(* Logix 5000 project; controller TFF vendor 1 type 14 code 107 rev 34.11; software revision 34.03; part 33 of 36 *)
(* tags used below, declared in another part *)
   Address : DINT;   // Temp Address
   Index : DINT;   // Index
   FlowPath : FlowPath[64];   // Flow Path Array
   PipeAnimation : PipeAnimation;   // HMI Pipe Animation Array
   PipeStatValueHMI : INT[224];   // Pipe Animation Value For HMI
   Rack_Murr_Node0_Smart : IO_Station;   // Status of Node 0 Smart
   Rack_Murr_Node1_TF2S : IO_Station;   // Status of Node 1 TF2S
   Rack_Murr_Node1_TF3S : IO_Station;   // Status of Node 1 TF3S
   Rack_Murr_Node3_PUMP : IO_Station;   // Status of Node 3 Pump
   Rack_Murr_Node4_Instrum_TFF1 : IO_Station;   // Status of Node 4 Instrum TFF1
   Rack_Murr_Node4_Instrum_TFF2 : IO_Station;   // Status of Node 4 Instrum TFF2
   Rack_Murr_Node4_Instrum_TFF3 : IO_Station;   // Status of Node 4 Instrum TFF3
   Rack_Murr_Node4_Instrum_TFF4 : IO_Station;   // Status of Node 4 Instrum TFF4
   Rack_Murr_Node4_Instrum_TFF5 : IO_Station;   // Status of Node 4 Instrum TFF5
   Rack_Murr_Node5_Tank100 : IO_Station;   // Status of Node 5 Tank 100L
   Rack_Murr_Node5_Tank250 : IO_Station;   // Status of Node 5 Tank 250L
   Rack_Murr_Node5_Tank50 : IO_Station;   // Status of Node 5 Tank 50L
   Rack_Murr_Node6_IND331_WI001 : IO_Station;   // Status of Node 6 IND331 WI001
   Rack_Murr_Node7_IND131_WI101 : IO_Station;   // Status of Node 7 IND131 WI101
   SIC001 : ALIAS FOR Drive[1];   // Feed Pump
   SIC002 : ALIAS FOR Drive[2];   // Transfer Pump
   Tank : TankManagement;   // Tank Management
   WI001 : ALIAS FOR AnalogPoint[15];   // Feed Bag Weight
   WI101 : ALIAS FOR AnalogPoint[0];   // Filtrate Weight
(* Process, continued *)

ROUTINE PipeAnimationHMI   (* ladder *)
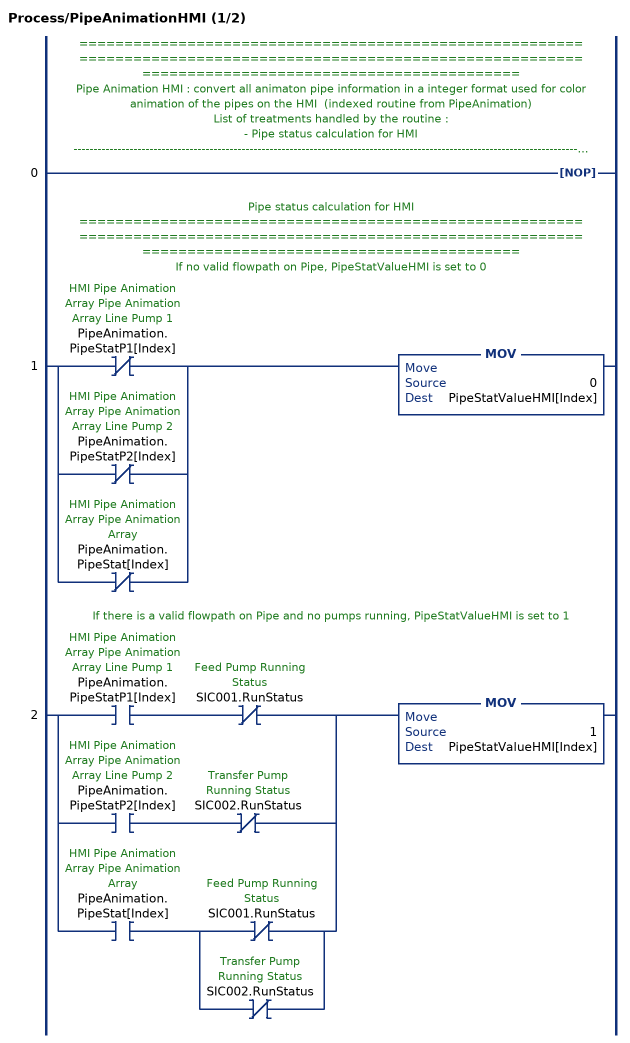
   // ==========================================================================================================================================================
   //                          Pipe Animation HMI : convert all animaton pipe information in a integer format used for color animation of the pipes on the HMI  (indexed routine from PipeAnimation)
   //                                                     List of treatments handled by the routine :
   //                                                          - Pipe status calculation for HMI
   //                                                     -----------------------------------------------------------------------------------------------------------------------------------------------------
   //                                                     History
   //                                                          2019-AUG-13 - Actemium - B. Roch - Initial version for Candidate Release 3.00.00.00.a
   // ========================================================================================================================================================
   0: NOP();
   // Pipe status calculation for HMI
   // ==========================================================================================================================================================
   // If no valid flowpath on Pipe, PipeStatValueHMI is set to 0
   1: [XIO(PipeAnimation.PipeStatP1[Index]) ,XIO(PipeAnimation.PipeStatP2[Index]) ,XIO(PipeAnimation.PipeStat[Index]) ]MOV(0,PipeStatValueHMI[Index]);
   // If there is a valid flowpath on Pipe and no pumps running, PipeStatValueHMI is set to 1
   2: [XIC(PipeAnimation.PipeStatP1[Index]) XIO(SIC001.RunStatus) ,XIC(PipeAnimation.PipeStatP2[Index]) XIO(SIC002.RunStatus) ,XIC(PipeAnimation.PipeStat[Index]) [XIO(SIC001.RunStatus) ,XIO(SIC002.RunStatus) ] ]MOV(1,PipeStatValueHMI[Index]);
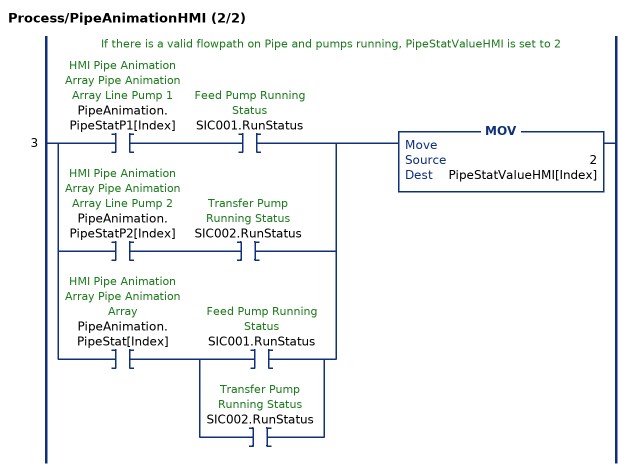
   // If there is a valid flowpath on Pipe and pumps running, PipeStatValueHMI is set to 2
   3: [XIC(PipeAnimation.PipeStatP1[Index]) XIC(SIC001.RunStatus) ,XIC(PipeAnimation.PipeStatP2[Index]) XIC(SIC002.RunStatus) ,XIC(PipeAnimation.PipeStat[Index]) [XIC(SIC001.RunStatus) ,XIC(SIC002.RunStatus) ] ]MOV(2,PipeStatValueHMI[Index]);
END_ROUTINE

ROUTINE Scale   (* function block diagram *)
// Scale Routine
   SHEET 1
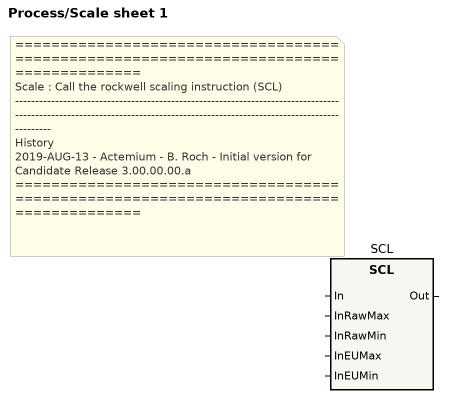
   // ======================================================================================
   // Scale : Call the rockwell scaling instruction (SCL)
   // ------------------------------------------------------------------------------------------------------------------------------------------------------------------
   // ---------
   // History
   //    2019-AUG-13 - Actemium - B. Roch - Initial version for Candidate Release 3.00.00.00.a
   // ======================================================================================
   SCL : SCL();   // unwired pins: In InRawMax InRawMin InEUMax InEUMin Out
END_ROUTINE

ROUTINE Station_Status   (* ladder *)
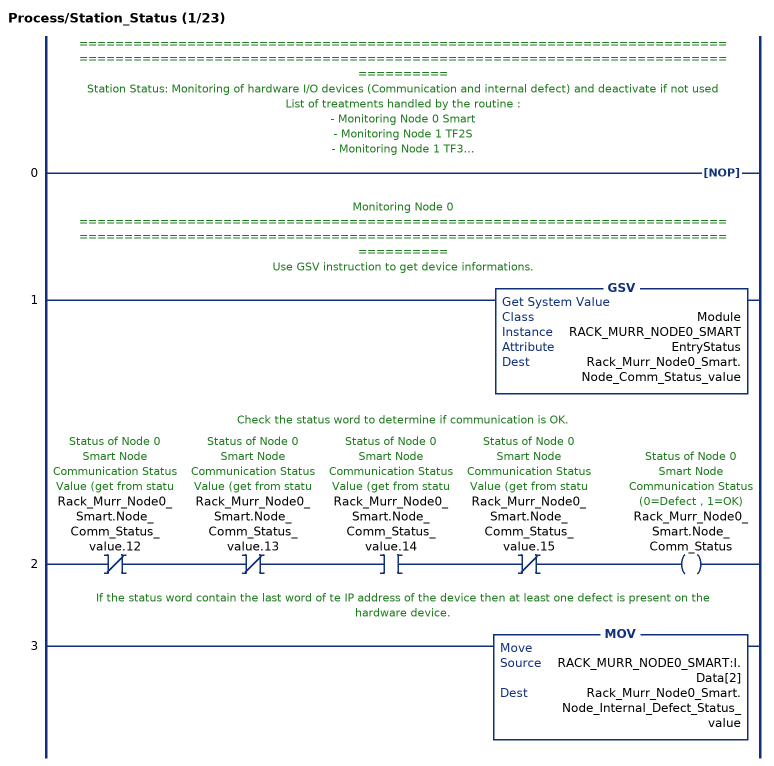
   // ==========================================================================================================================================================
   //                                                                   Station Status: Monitoring of hardware I/O devices (Communication and internal defect) and deactivate if not used
   //                                                     List of treatments handled by the routine :
   //                                                        - Monitoring Node 0 Smart
   //                                                        - Monitoring Node 1 TF2S
   //                                                        - Monitoring Node 1 TF3S
   //                                                        - Monitoring Node 3 PUMP
   //                                                        - Monitoring Node 4 INTRUM TFF1
   //                                                        - Monitoring Node 4 INTRUM TFF2
   //                                                        - Monitoring Node 4 INTRUM TFF3
   //                                                        - Monitoring Node 4 INTRUM TFF4
   //                                                        - Monitoring Node 4 INTRUM TFF5
   //                                                        - Monitoring Node 5 TANK50
   //                                                        - Monitoring Node 5 TANK100
   //                                                        - Monitoring Node 5 TANK250
   //                                                        - Monitoring Node 6 IND331 WI001
   //                                                        - Monitoring Node 7 IND131 WI101
   //                                                        - Deactivate / Activate devices
   //                                                     -----------------------------------------------------------------------------------------------------------------------------------------------------
   //                                                     History
   //                                                          2019-AUG-13 - Actemium - B. Roch - Initial version for Candidate Release 3.00.00.00.a
   // ========================================================================================================================================================
   0: NOP();
   // Monitoring Node 0
   // ==========================================================================================================================================================
   // Use GSV instruction to get device informations.
   1: GSV(Module,RACK_MURR_NODE0_SMART,EntryStatus,Rack_Murr_Node0_Smart.Node_Comm_Status_value);
   // Check the status word to determine if communication is OK.
   2: XIO(Rack_Murr_Node0_Smart.Node_Comm_Status_value.12)XIO(Rack_Murr_Node0_Smart.Node_Comm_Status_value.13)XIC(Rack_Murr_Node0_Smart.Node_Comm_Status_value.14)XIO(Rack_Murr_Node0_Smart.Node_Comm_Status_value.15)OTE(Rack_Murr_Node0_Smart.Node_Comm_Status);
   // If the status word contain the last word of te IP address of the device then at least one defect is present on the hardware device.
   3: MOV(RACK_MURR_NODE0_SMART:I.Data[2],Rack_Murr_Node0_Smart.Node_Internal_Defect_Status_value);
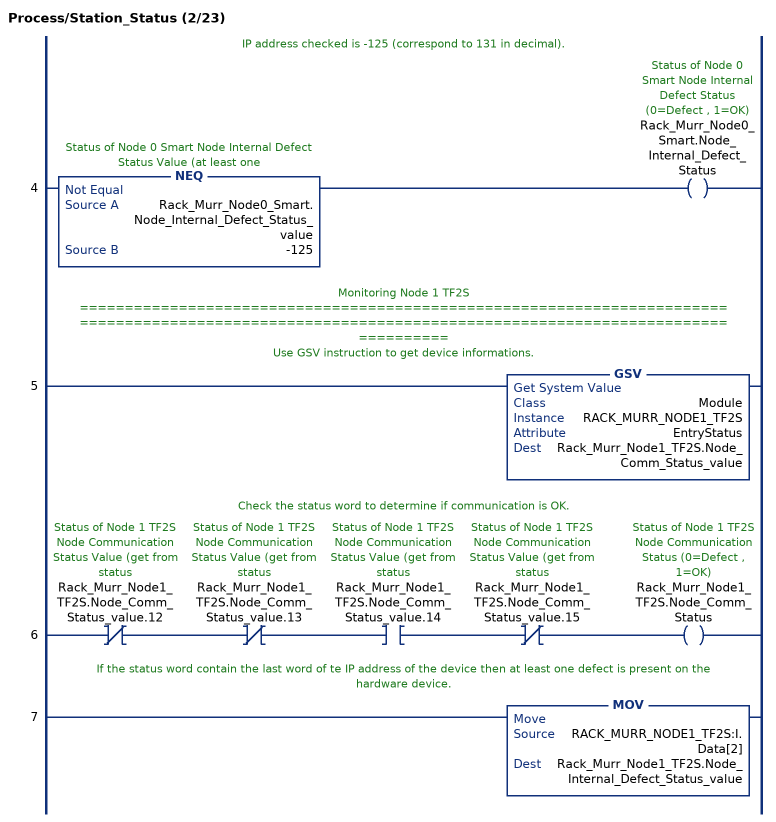
   // IP address checked is -125 (correspond to 131 in decimal).
   4: NEQ(Rack_Murr_Node0_Smart.Node_Internal_Defect_Status_value,-125)OTE(Rack_Murr_Node0_Smart.Node_Internal_Defect_Status);
   // Monitoring Node 1 TF2S
   // ==========================================================================================================================================================
   // Use GSV instruction to get device informations.
   5: GSV(Module,RACK_MURR_NODE1_TF2S,EntryStatus,Rack_Murr_Node1_TF2S.Node_Comm_Status_value);
   // Check the status word to determine if communication is OK.
   6: XIO(Rack_Murr_Node1_TF2S.Node_Comm_Status_value.12)XIO(Rack_Murr_Node1_TF2S.Node_Comm_Status_value.13)XIC(Rack_Murr_Node1_TF2S.Node_Comm_Status_value.14)XIO(Rack_Murr_Node1_TF2S.Node_Comm_Status_value.15)OTE(Rack_Murr_Node1_TF2S.Node_Comm_Status);
   // If the status word contain the last word of te IP address of the device then at least one defect is present on the hardware device.
   7: MOV(RACK_MURR_NODE1_TF2S:I.Data[2],Rack_Murr_Node1_TF2S.Node_Internal_Defect_Status_value);
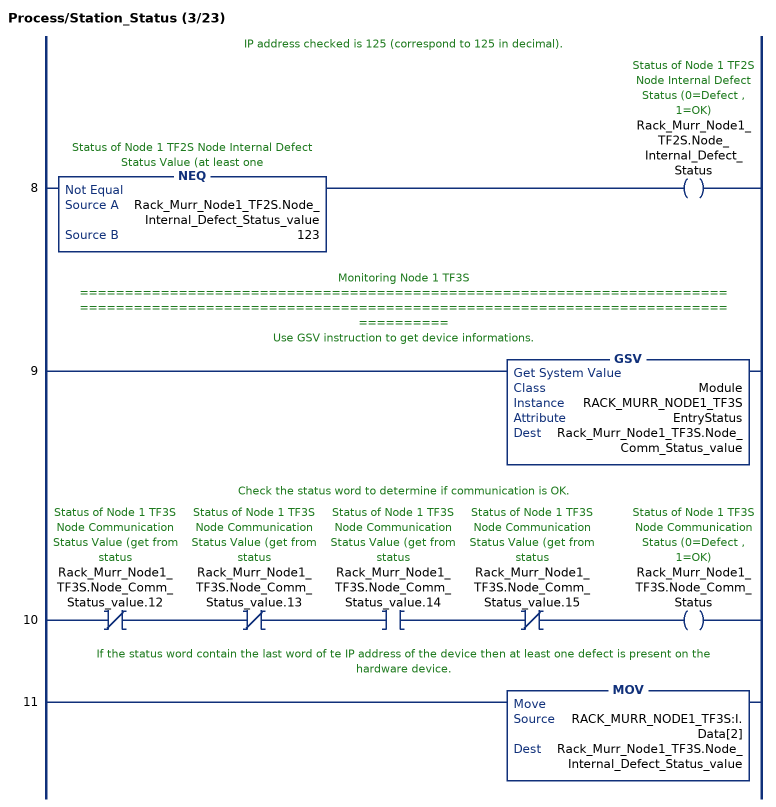
   // IP address checked is 125 (correspond to 125 in decimal).
   8: NEQ(Rack_Murr_Node1_TF2S.Node_Internal_Defect_Status_value,123)OTE(Rack_Murr_Node1_TF2S.Node_Internal_Defect_Status);
   // Monitoring Node 1 TF3S
   // ==========================================================================================================================================================
   // Use GSV instruction to get device informations.
   9: GSV(Module,RACK_MURR_NODE1_TF3S,EntryStatus,Rack_Murr_Node1_TF3S.Node_Comm_Status_value);
   // Check the status word to determine if communication is OK.
   10: XIO(Rack_Murr_Node1_TF3S.Node_Comm_Status_value.12)XIO(Rack_Murr_Node1_TF3S.Node_Comm_Status_value.13)XIC(Rack_Murr_Node1_TF3S.Node_Comm_Status_value.14)XIO(Rack_Murr_Node1_TF3S.Node_Comm_Status_value.15)OTE(Rack_Murr_Node1_TF3S.Node_Comm_Status);
   // If the status word contain the last word of te IP address of the device then at least one defect is present on the hardware device.
   11: MOV(RACK_MURR_NODE1_TF3S:I.Data[2],Rack_Murr_Node1_TF3S.Node_Internal_Defect_Status_value);
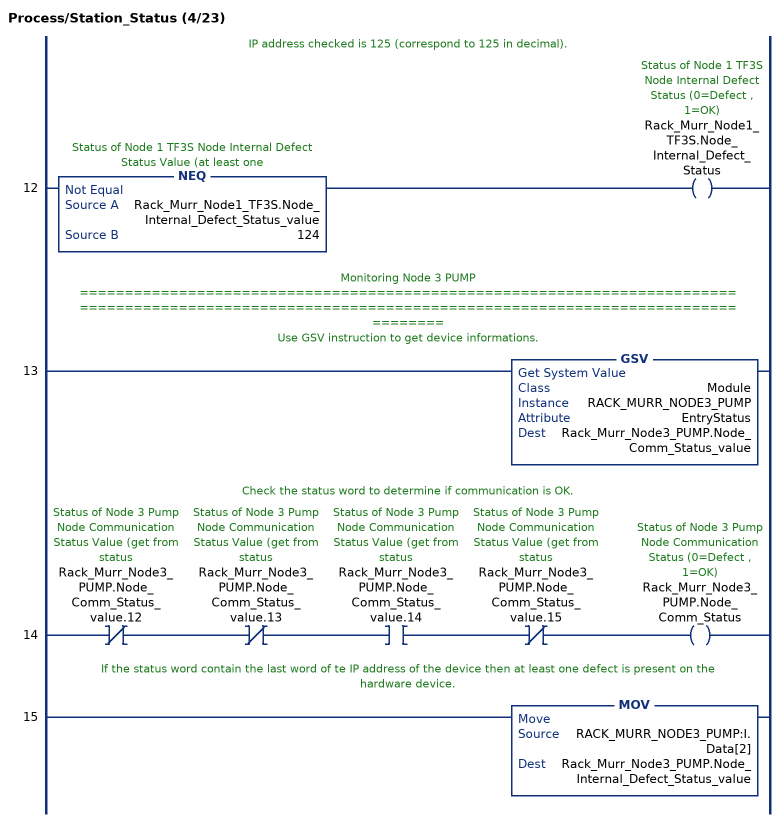
   // IP address checked is 125 (correspond to 125 in decimal).
   12: NEQ(Rack_Murr_Node1_TF3S.Node_Internal_Defect_Status_value,124)OTE(Rack_Murr_Node1_TF3S.Node_Internal_Defect_Status);
   // Monitoring Node 3 PUMP
   // ==========================================================================================================================================================
   // Use GSV instruction to get device informations.
   13: GSV(Module,RACK_MURR_NODE3_PUMP,EntryStatus,Rack_Murr_Node3_PUMP.Node_Comm_Status_value);
   // Check the status word to determine if communication is OK.
   14: XIO(Rack_Murr_Node3_PUMP.Node_Comm_Status_value.12)XIO(Rack_Murr_Node3_PUMP.Node_Comm_Status_value.13)XIC(Rack_Murr_Node3_PUMP.Node_Comm_Status_value.14)XIO(Rack_Murr_Node3_PUMP.Node_Comm_Status_value.15)OTE(Rack_Murr_Node3_PUMP.Node_Comm_Status);
   // If the status word contain the last word of te IP address of the device then at least one defect is present on the hardware device.
   15: MOV(RACK_MURR_NODE3_PUMP:I.Data[2],Rack_Murr_Node3_PUMP.Node_Internal_Defect_Status_value);
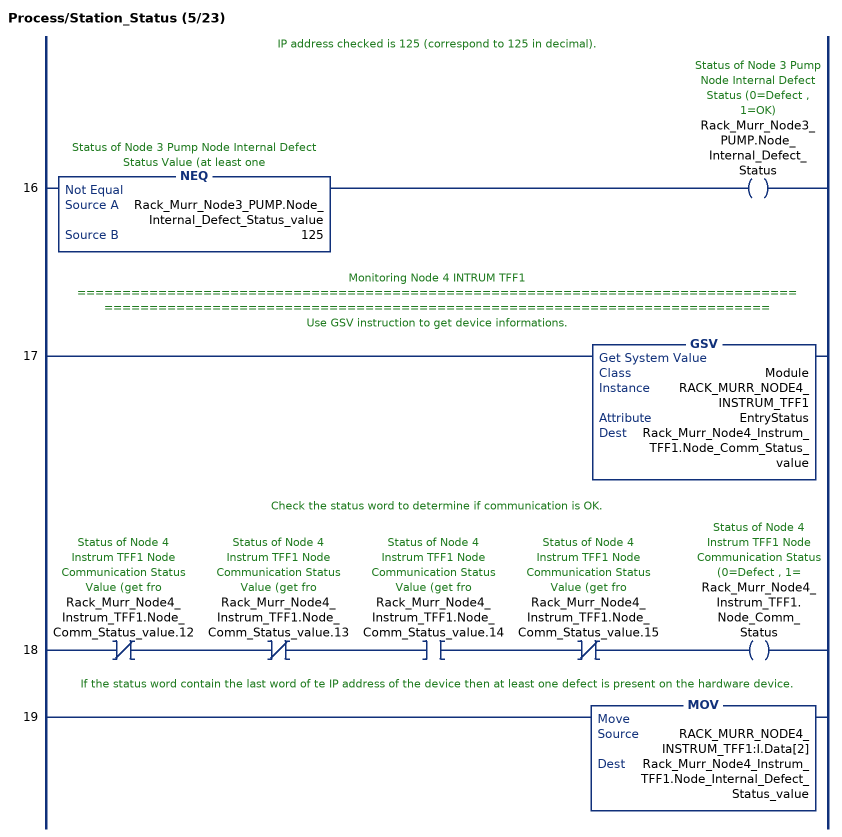
   // IP address checked is 125 (correspond to 125 in decimal).
   16: NEQ(Rack_Murr_Node3_PUMP.Node_Internal_Defect_Status_value,125)OTE(Rack_Murr_Node3_PUMP.Node_Internal_Defect_Status);
   // Monitoring Node 4 INTRUM TFF1
   // ==========================================================================================================================================================
   // Use GSV instruction to get device informations.
   17: GSV(Module,RACK_MURR_NODE4_INSTRUM_TFF1,EntryStatus,Rack_Murr_Node4_Instrum_TFF1.Node_Comm_Status_value);
   // Check the status word to determine if communication is OK.
   18: XIO(Rack_Murr_Node4_Instrum_TFF1.Node_Comm_Status_value.12)XIO(Rack_Murr_Node4_Instrum_TFF1.Node_Comm_Status_value.13)XIC(Rack_Murr_Node4_Instrum_TFF1.Node_Comm_Status_value.14)XIO(Rack_Murr_Node4_Instrum_TFF1.Node_Comm_Status_value.15)OTE(Rack_Murr_Node4_Instrum_TFF1.Node_Comm_Status);
   // If the status word contain the last word of te IP address of the device then at least one defect is present on the hardware device.
   19: MOV(RACK_MURR_NODE4_INSTRUM_TFF1:I.Data[2],Rack_Murr_Node4_Instrum_TFF1.Node_Internal_Defect_Status_value);
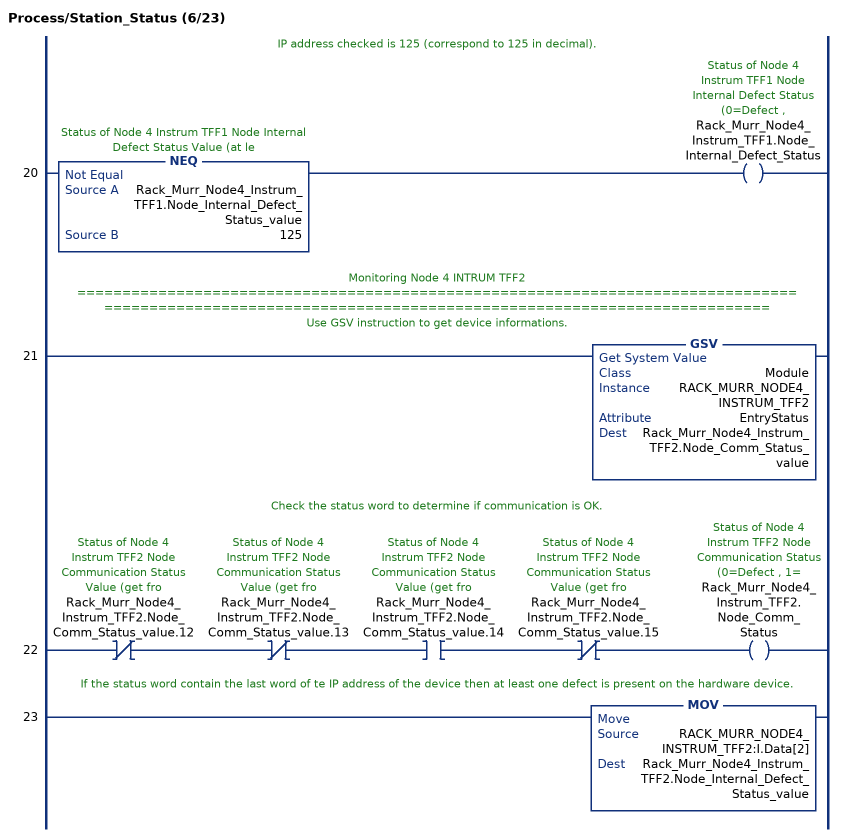
   // IP address checked is 125 (correspond to 125 in decimal).
   20: NEQ(Rack_Murr_Node4_Instrum_TFF1.Node_Internal_Defect_Status_value,125)OTE(Rack_Murr_Node4_Instrum_TFF1.Node_Internal_Defect_Status);
   // Monitoring Node 4 INTRUM TFF2
   // ==========================================================================================================================================================
   // Use GSV instruction to get device informations.
   21: GSV(Module,RACK_MURR_NODE4_INSTRUM_TFF2,EntryStatus,Rack_Murr_Node4_Instrum_TFF2.Node_Comm_Status_value);
   // Check the status word to determine if communication is OK.
   22: XIO(Rack_Murr_Node4_Instrum_TFF2.Node_Comm_Status_value.12)XIO(Rack_Murr_Node4_Instrum_TFF2.Node_Comm_Status_value.13)XIC(Rack_Murr_Node4_Instrum_TFF2.Node_Comm_Status_value.14)XIO(Rack_Murr_Node4_Instrum_TFF2.Node_Comm_Status_value.15)OTE(Rack_Murr_Node4_Instrum_TFF2.Node_Comm_Status);
   // If the status word contain the last word of te IP address of the device then at least one defect is present on the hardware device.
   23: MOV(RACK_MURR_NODE4_INSTRUM_TFF2:I.Data[2],Rack_Murr_Node4_Instrum_TFF2.Node_Internal_Defect_Status_value);
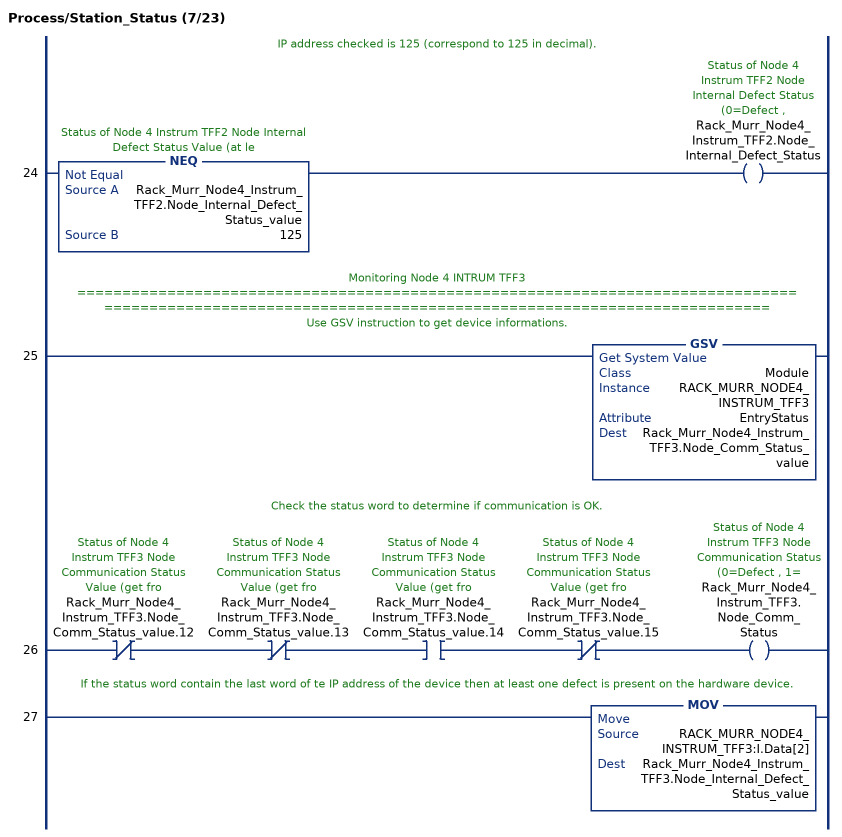
   // IP address checked is 125 (correspond to 125 in decimal).
   24: NEQ(Rack_Murr_Node4_Instrum_TFF2.Node_Internal_Defect_Status_value,125)OTE(Rack_Murr_Node4_Instrum_TFF2.Node_Internal_Defect_Status);
   // Monitoring Node 4 INTRUM TFF3
   // ==========================================================================================================================================================
   // Use GSV instruction to get device informations.
   25: GSV(Module,RACK_MURR_NODE4_INSTRUM_TFF3,EntryStatus,Rack_Murr_Node4_Instrum_TFF3.Node_Comm_Status_value);
   // Check the status word to determine if communication is OK.
   26: XIO(Rack_Murr_Node4_Instrum_TFF3.Node_Comm_Status_value.12)XIO(Rack_Murr_Node4_Instrum_TFF3.Node_Comm_Status_value.13)XIC(Rack_Murr_Node4_Instrum_TFF3.Node_Comm_Status_value.14)XIO(Rack_Murr_Node4_Instrum_TFF3.Node_Comm_Status_value.15)OTE(Rack_Murr_Node4_Instrum_TFF3.Node_Comm_Status);
   // If the status word contain the last word of te IP address of the device then at least one defect is present on the hardware device.
   27: MOV(RACK_MURR_NODE4_INSTRUM_TFF3:I.Data[2],Rack_Murr_Node4_Instrum_TFF3.Node_Internal_Defect_Status_value);
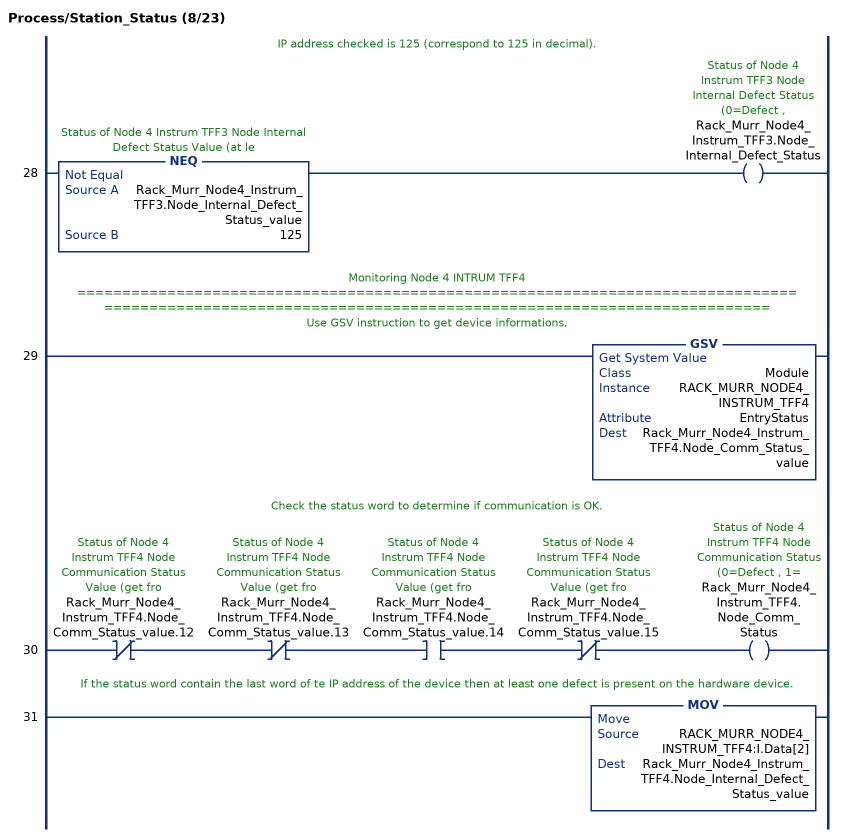
   // IP address checked is 125 (correspond to 125 in decimal).
   28: NEQ(Rack_Murr_Node4_Instrum_TFF3.Node_Internal_Defect_Status_value,125)OTE(Rack_Murr_Node4_Instrum_TFF3.Node_Internal_Defect_Status);
   // Monitoring Node 4 INTRUM TFF4
   // ==========================================================================================================================================================
   // Use GSV instruction to get device informations.
   29: GSV(Module,RACK_MURR_NODE4_INSTRUM_TFF4,EntryStatus,Rack_Murr_Node4_Instrum_TFF4.Node_Comm_Status_value);
   // Check the status word to determine if communication is OK.
   30: XIO(Rack_Murr_Node4_Instrum_TFF4.Node_Comm_Status_value.12)XIO(Rack_Murr_Node4_Instrum_TFF4.Node_Comm_Status_value.13)XIC(Rack_Murr_Node4_Instrum_TFF4.Node_Comm_Status_value.14)XIO(Rack_Murr_Node4_Instrum_TFF4.Node_Comm_Status_value.15)OTE(Rack_Murr_Node4_Instrum_TFF4.Node_Comm_Status);
   // If the status word contain the last word of te IP address of the device then at least one defect is present on the hardware device.
   31: MOV(RACK_MURR_NODE4_INSTRUM_TFF4:I.Data[2],Rack_Murr_Node4_Instrum_TFF4.Node_Internal_Defect_Status_value);
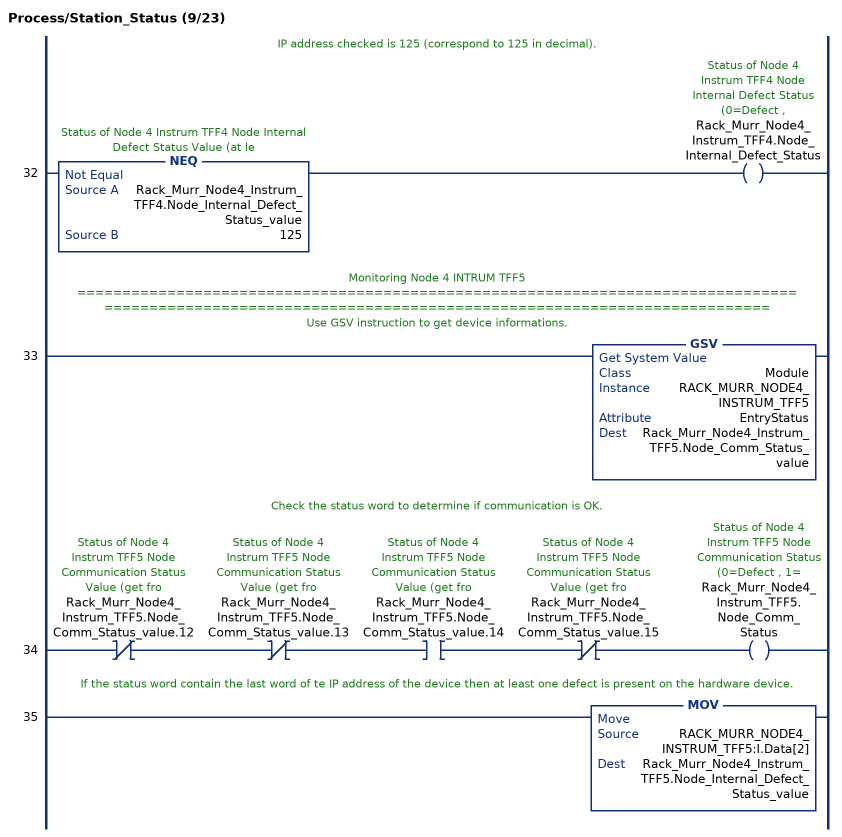
   // IP address checked is 125 (correspond to 125 in decimal).
   32: NEQ(Rack_Murr_Node4_Instrum_TFF4.Node_Internal_Defect_Status_value,125)OTE(Rack_Murr_Node4_Instrum_TFF4.Node_Internal_Defect_Status);
   // Monitoring Node 4 INTRUM TFF5
   // ==========================================================================================================================================================
   // Use GSV instruction to get device informations.
   33: GSV(Module,RACK_MURR_NODE4_INSTRUM_TFF5,EntryStatus,Rack_Murr_Node4_Instrum_TFF5.Node_Comm_Status_value);
   // Check the status word to determine if communication is OK.
   34: XIO(Rack_Murr_Node4_Instrum_TFF5.Node_Comm_Status_value.12)XIO(Rack_Murr_Node4_Instrum_TFF5.Node_Comm_Status_value.13)XIC(Rack_Murr_Node4_Instrum_TFF5.Node_Comm_Status_value.14)XIO(Rack_Murr_Node4_Instrum_TFF5.Node_Comm_Status_value.15)OTE(Rack_Murr_Node4_Instrum_TFF5.Node_Comm_Status);
   // If the status word contain the last word of te IP address of the device then at least one defect is present on the hardware device.
   35: MOV(RACK_MURR_NODE4_INSTRUM_TFF5:I.Data[2],Rack_Murr_Node4_Instrum_TFF5.Node_Internal_Defect_Status_value);
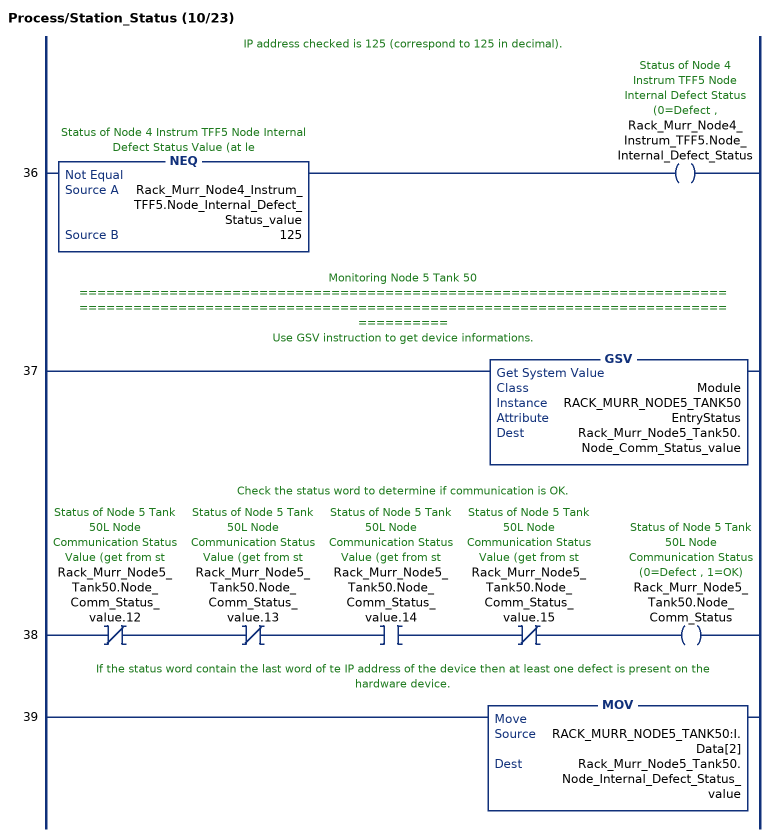
   // IP address checked is 125 (correspond to 125 in decimal).
   36: NEQ(Rack_Murr_Node4_Instrum_TFF5.Node_Internal_Defect_Status_value,125)OTE(Rack_Murr_Node4_Instrum_TFF5.Node_Internal_Defect_Status);
   // Monitoring Node 5 Tank 50
   // ==========================================================================================================================================================
   // Use GSV instruction to get device informations.
   37: GSV(Module,RACK_MURR_NODE5_TANK50,EntryStatus,Rack_Murr_Node5_Tank50.Node_Comm_Status_value);
   // Check the status word to determine if communication is OK.
   38: XIO(Rack_Murr_Node5_Tank50.Node_Comm_Status_value.12)XIO(Rack_Murr_Node5_Tank50.Node_Comm_Status_value.13)XIC(Rack_Murr_Node5_Tank50.Node_Comm_Status_value.14)XIO(Rack_Murr_Node5_Tank50.Node_Comm_Status_value.15)OTE(Rack_Murr_Node5_Tank50.Node_Comm_Status);
   // If the status word contain the last word of te IP address of the device then at least one defect is present on the hardware device.
   39: MOV(RACK_MURR_NODE5_TANK50:I.Data[2],Rack_Murr_Node5_Tank50.Node_Internal_Defect_Status_value);
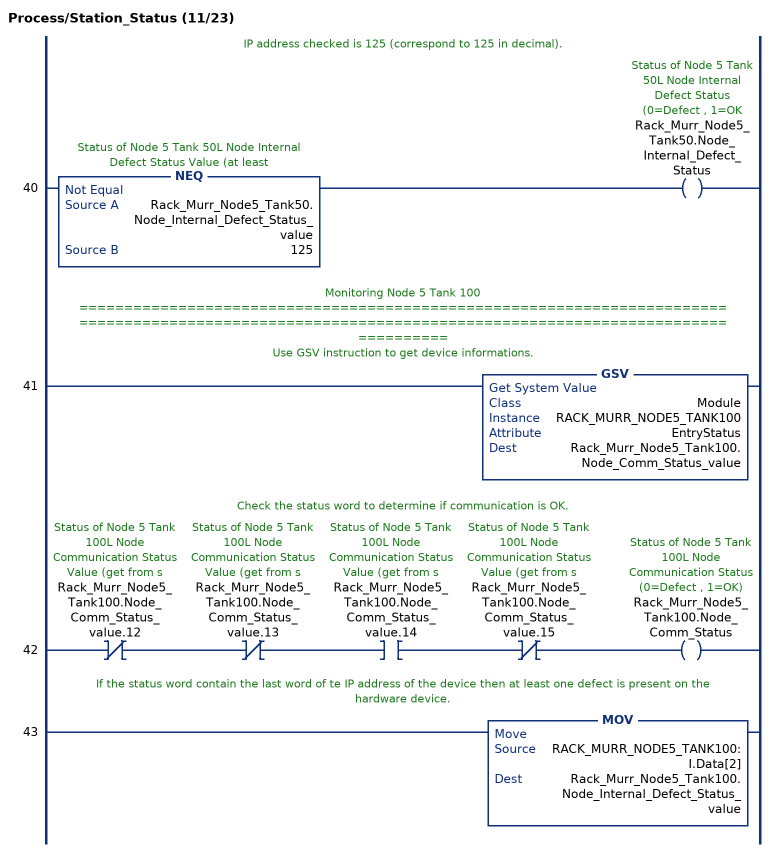
   // IP address checked is 125 (correspond to 125 in decimal).
   40: NEQ(Rack_Murr_Node5_Tank50.Node_Internal_Defect_Status_value,125)OTE(Rack_Murr_Node5_Tank50.Node_Internal_Defect_Status);
   // Monitoring Node 5 Tank 100
   // ==========================================================================================================================================================
   // Use GSV instruction to get device informations.
   41: GSV(Module,RACK_MURR_NODE5_TANK100,EntryStatus,Rack_Murr_Node5_Tank100.Node_Comm_Status_value);
   // Check the status word to determine if communication is OK.
   42: XIO(Rack_Murr_Node5_Tank100.Node_Comm_Status_value.12)XIO(Rack_Murr_Node5_Tank100.Node_Comm_Status_value.13)XIC(Rack_Murr_Node5_Tank100.Node_Comm_Status_value.14)XIO(Rack_Murr_Node5_Tank100.Node_Comm_Status_value.15)OTE(Rack_Murr_Node5_Tank100.Node_Comm_Status);
   // If the status word contain the last word of te IP address of the device then at least one defect is present on the hardware device.
   43: MOV(RACK_MURR_NODE5_TANK100:I.Data[2],Rack_Murr_Node5_Tank100.Node_Internal_Defect_Status_value);
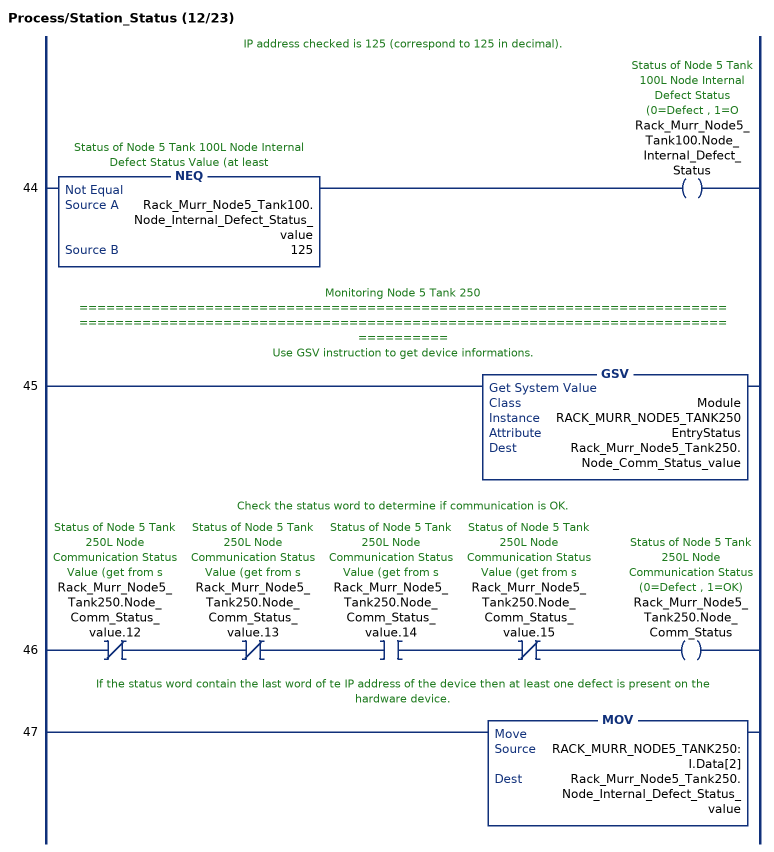
   // IP address checked is 125 (correspond to 125 in decimal).
   44: NEQ(Rack_Murr_Node5_Tank100.Node_Internal_Defect_Status_value,125)OTE(Rack_Murr_Node5_Tank100.Node_Internal_Defect_Status);
   // Monitoring Node 5 Tank 250
   // ==========================================================================================================================================================
   // Use GSV instruction to get device informations.
   45: GSV(Module,RACK_MURR_NODE5_TANK250,EntryStatus,Rack_Murr_Node5_Tank250.Node_Comm_Status_value);
   // Check the status word to determine if communication is OK.
   46: XIO(Rack_Murr_Node5_Tank250.Node_Comm_Status_value.12)XIO(Rack_Murr_Node5_Tank250.Node_Comm_Status_value.13)XIC(Rack_Murr_Node5_Tank250.Node_Comm_Status_value.14)XIO(Rack_Murr_Node5_Tank250.Node_Comm_Status_value.15)OTE(Rack_Murr_Node5_Tank250.Node_Comm_Status);
   // If the status word contain the last word of te IP address of the device then at least one defect is present on the hardware device.
   47: MOV(RACK_MURR_NODE5_TANK250:I.Data[2],Rack_Murr_Node5_Tank250.Node_Internal_Defect_Status_value);
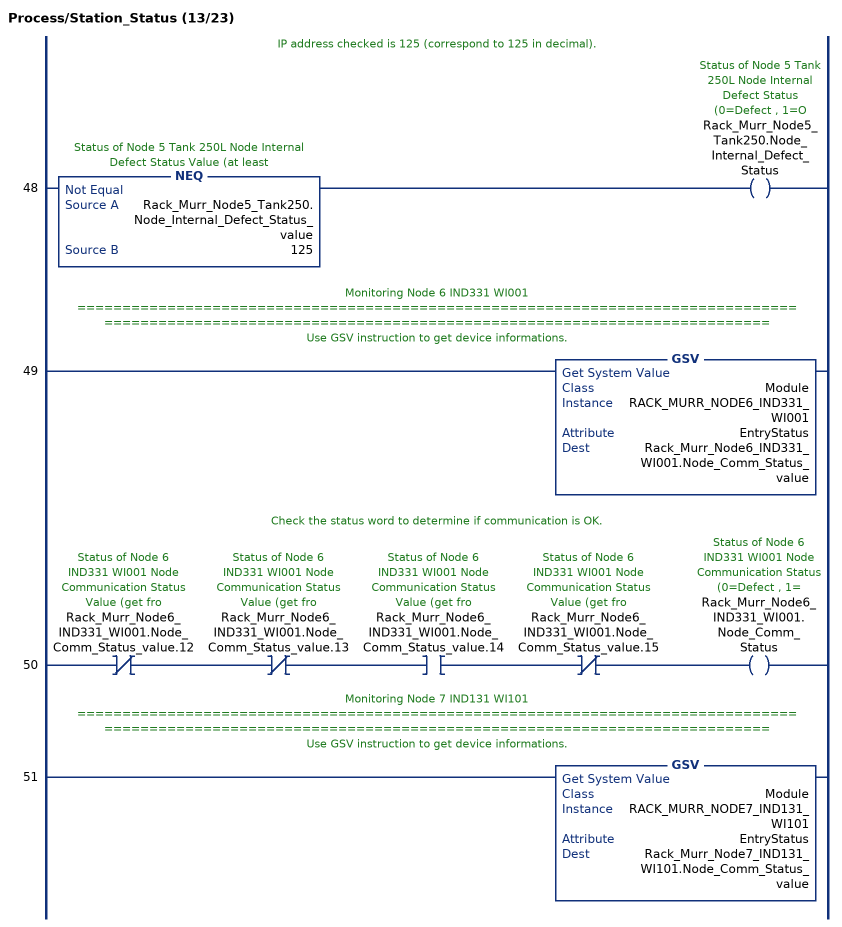
   // IP address checked is 125 (correspond to 125 in decimal).
   48: NEQ(Rack_Murr_Node5_Tank250.Node_Internal_Defect_Status_value,125)OTE(Rack_Murr_Node5_Tank250.Node_Internal_Defect_Status);
   // Monitoring Node 6 IND331 WI001
   // ==========================================================================================================================================================
   // Use GSV instruction to get device informations.
   49: GSV(Module,RACK_MURR_NODE6_IND331_WI001,EntryStatus,Rack_Murr_Node6_IND331_WI001.Node_Comm_Status_value);
   // Check the status word to determine if communication is OK.
   50: XIO(Rack_Murr_Node6_IND331_WI001.Node_Comm_Status_value.12)XIO(Rack_Murr_Node6_IND331_WI001.Node_Comm_Status_value.13)XIC(Rack_Murr_Node6_IND331_WI001.Node_Comm_Status_value.14)XIO(Rack_Murr_Node6_IND331_WI001.Node_Comm_Status_value.15)OTE(Rack_Murr_Node6_IND331_WI001.Node_Comm_Status);
   // Monitoring Node 7 IND131 WI101
   // ==========================================================================================================================================================
   // Use GSV instruction to get device informations.
   51: GSV(Module,RACK_MURR_NODE7_IND131_WI101,EntryStatus,Rack_Murr_Node7_IND131_WI101.Node_Comm_Status_value);
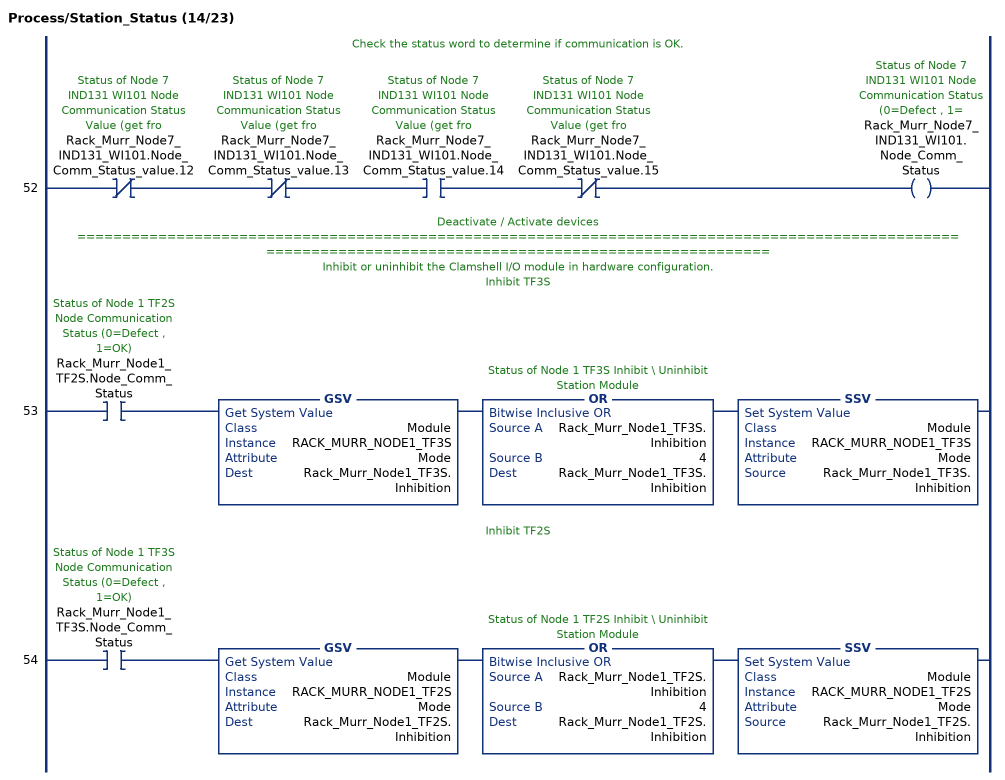
   // Check the status word to determine if communication is OK.
   52: XIO(Rack_Murr_Node7_IND131_WI101.Node_Comm_Status_value.12)XIO(Rack_Murr_Node7_IND131_WI101.Node_Comm_Status_value.13)XIC(Rack_Murr_Node7_IND131_WI101.Node_Comm_Status_value.14)XIO(Rack_Murr_Node7_IND131_WI101.Node_Comm_Status_value.15)OTE(Rack_Murr_Node7_IND131_WI101.Node_Comm_Status);
   // Deactivate / Activate devices
   // ==========================================================================================================================================================
   // Inhibit or uninhibit the Clamshell I/O module in hardware configuration.
   // Inhibit TF3S
   53: XIC(Rack_Murr_Node1_TF2S.Node_Comm_Status)GSV(Module,RACK_MURR_NODE1_TF3S,Mode,Rack_Murr_Node1_TF3S.Inhibition)OR(Rack_Murr_Node1_TF3S.Inhibition,4,Rack_Murr_Node1_TF3S.Inhibition)SSV(Module,RACK_MURR_NODE1_TF3S,Mode,Rack_Murr_Node1_TF3S.Inhibition);
   // Inhibit TF2S
   54: XIC(Rack_Murr_Node1_TF3S.Node_Comm_Status)GSV(Module,RACK_MURR_NODE1_TF2S,Mode,Rack_Murr_Node1_TF2S.Inhibition)OR(Rack_Murr_Node1_TF2S.Inhibition,4,Rack_Murr_Node1_TF2S.Inhibition)SSV(Module,RACK_MURR_NODE1_TF2S,Mode,Rack_Murr_Node1_TF2S.Inhibition);
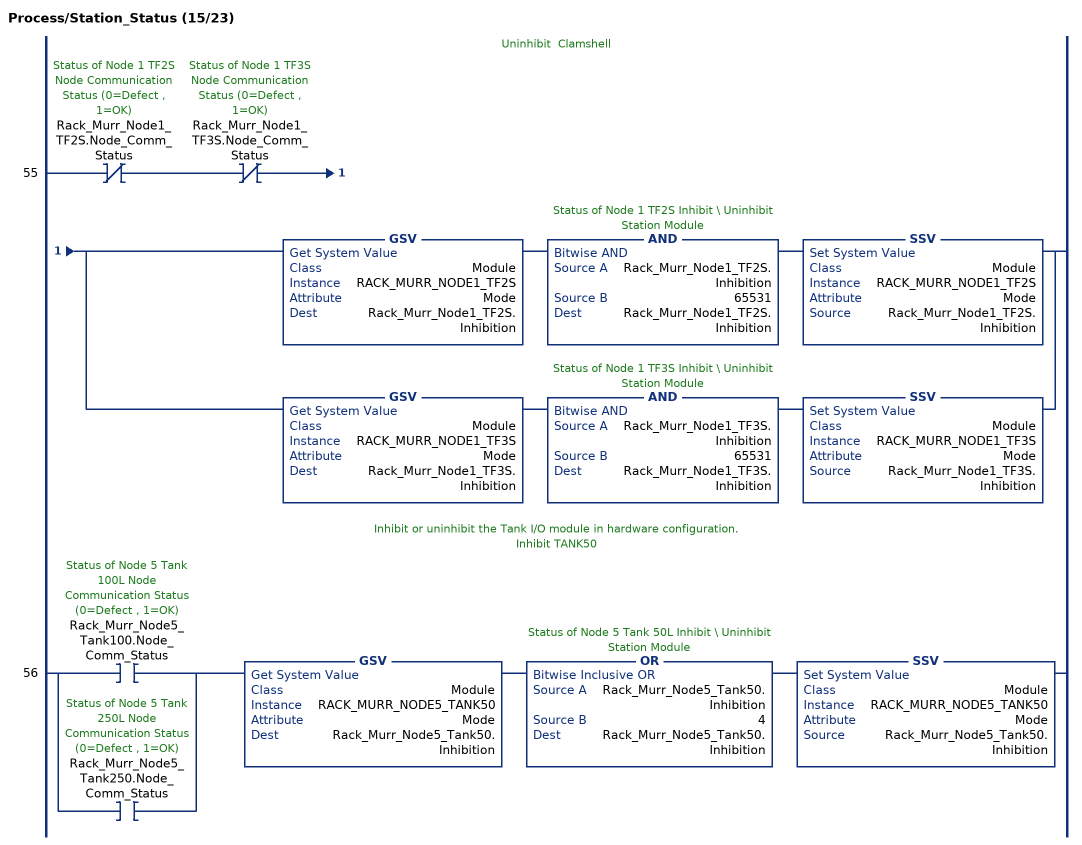
   // Uninhibit  Clamshell
   55: XIO(Rack_Murr_Node1_TF2S.Node_Comm_Status)XIO(Rack_Murr_Node1_TF3S.Node_Comm_Status)[GSV(Module,RACK_MURR_NODE1_TF2S,Mode,Rack_Murr_Node1_TF2S.Inhibition) AND(Rack_Murr_Node1_TF2S.Inhibition,65531,Rack_Murr_Node1_TF2S.Inhibition) SSV(Module,RACK_MURR_NODE1_TF2S,Mode,Rack_Murr_Node1_TF2S.Inhibition) ,GSV(Module,RACK_MURR_NODE1_TF3S,Mode,Rack_Murr_Node1_TF3S.Inhibition) AND(Rack_Murr_Node1_TF3S.Inhibition,65531,Rack_Murr_Node1_TF3S.Inhibition) SSV(Module,RACK_MURR_NODE1_TF3S,Mode,Rack_Murr_Node1_TF3S.Inhibition) ];
   // Inhibit or uninhibit the Tank I/O module in hardware configuration.
   // Inhibit TANK50
   56: [XIC(Rack_Murr_Node5_Tank100.Node_Comm_Status) ,XIC(Rack_Murr_Node5_Tank250.Node_Comm_Status) ]GSV(Module,RACK_MURR_NODE5_TANK50,Mode,Rack_Murr_Node5_Tank50.Inhibition)OR(Rack_Murr_Node5_Tank50.Inhibition,4,Rack_Murr_Node5_Tank50.Inhibition)SSV(Module,RACK_MURR_NODE5_TANK50,Mode,Rack_Murr_Node5_Tank50.Inhibition);
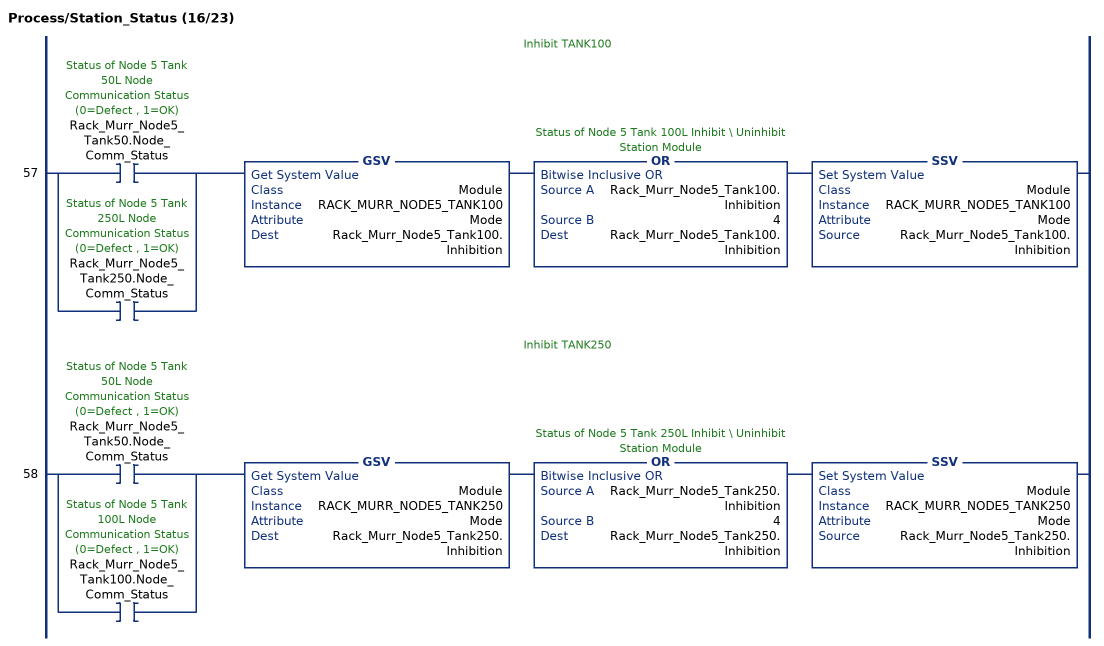
   // Inhibit TANK100
   57: [XIC(Rack_Murr_Node5_Tank50.Node_Comm_Status) ,XIC(Rack_Murr_Node5_Tank250.Node_Comm_Status) ]GSV(Module,RACK_MURR_NODE5_TANK100,Mode,Rack_Murr_Node5_Tank100.Inhibition)OR(Rack_Murr_Node5_Tank100.Inhibition,4,Rack_Murr_Node5_Tank100.Inhibition)SSV(Module,RACK_MURR_NODE5_TANK100,Mode,Rack_Murr_Node5_Tank100.Inhibition);
   // Inhibit TANK250
   58: [XIC(Rack_Murr_Node5_Tank50.Node_Comm_Status) ,XIC(Rack_Murr_Node5_Tank100.Node_Comm_Status) ]GSV(Module,RACK_MURR_NODE5_TANK250,Mode,Rack_Murr_Node5_Tank250.Inhibition)OR(Rack_Murr_Node5_Tank250.Inhibition,4,Rack_Murr_Node5_Tank250.Inhibition)SSV(Module,RACK_MURR_NODE5_TANK250,Mode,Rack_Murr_Node5_Tank250.Inhibition);
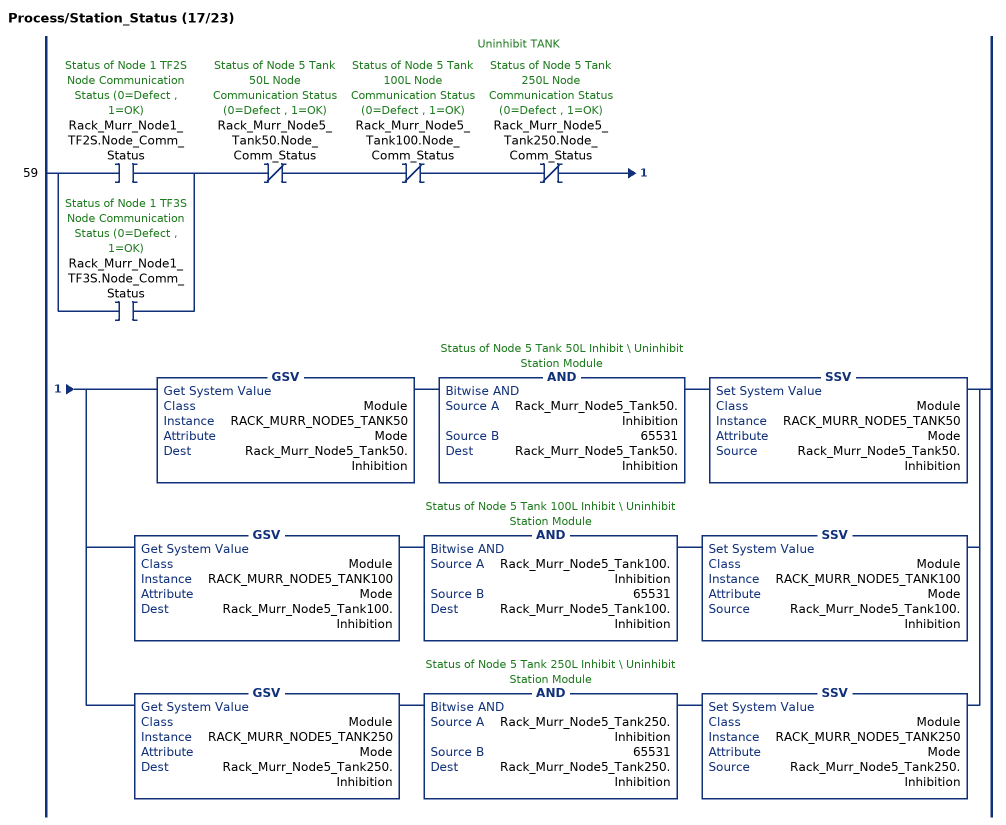
   // Uninhibit TANK
   59: [XIC(Rack_Murr_Node1_TF2S.Node_Comm_Status) ,XIC(Rack_Murr_Node1_TF3S.Node_Comm_Status) ]XIO(Rack_Murr_Node5_Tank50.Node_Comm_Status)XIO(Rack_Murr_Node5_Tank100.Node_Comm_Status)XIO(Rack_Murr_Node5_Tank250.Node_Comm_Status)[GSV(Module,RACK_MURR_NODE5_TANK50,Mode,Rack_Murr_Node5_Tank50.Inhibition) AND(Rack_Murr_Node5_Tank50.Inhibition,65531,Rack_Murr_Node5_Tank50.Inhibition) SSV(Module,RACK_MURR_NODE5_TANK50,Mode,Rack_Murr_Node5_Tank50.Inhibition) ,GSV(Module,RACK_MURR_NODE5_TANK100,Mode,Rack_Murr_Node5_Tank100.Inhibition) AND(Rack_Murr_Node5_Tank100.Inhibition,65531,Rack_Murr_Node5_Tank100.Inhibition) SSV(Module,RACK_MURR_NODE5_TANK100,Mode,Rack_Murr_Node5_Tank100.Inhibition) ,GSV(Module,RACK_MURR_NODE5_TANK250,Mode,Rack_Murr_Node5_Tank250.Inhibition) AND(Rack_Murr_Node5_Tank250.Inhibition,65531,Rack_Murr_Node5_Tank250.Inhibition) SSV(Module,RACK_MURR_NODE5_TANK250,Mode,Rack_Murr_Node5_Tank250.Inhibition) ];
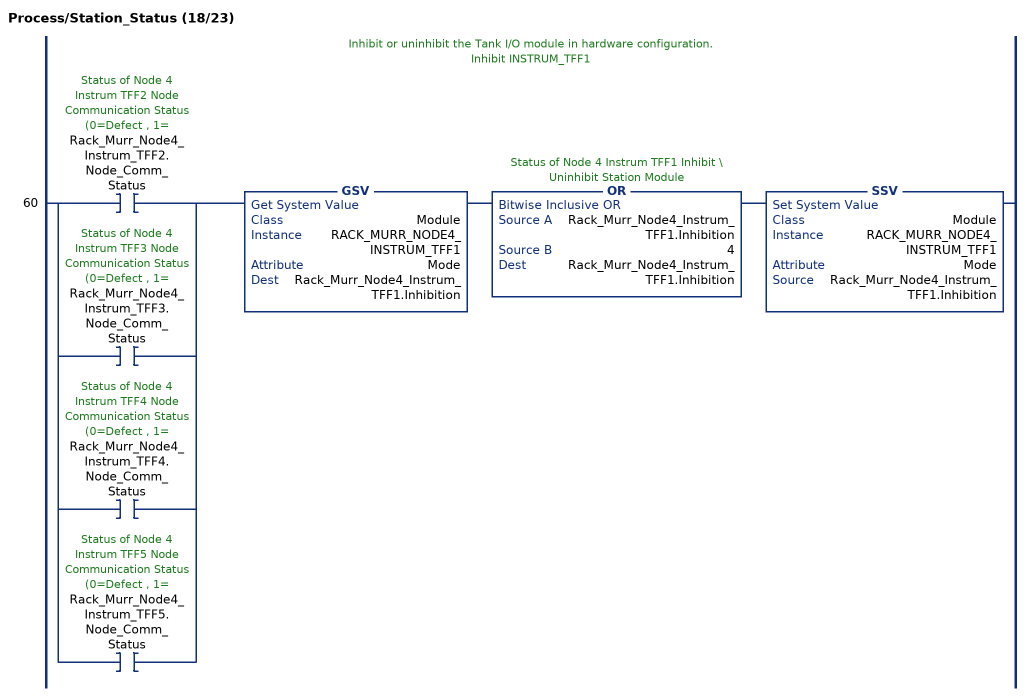
   // Inhibit or uninhibit the Tank I/O module in hardware configuration.
   // Inhibit INSTRUM_TFF1
   60: [XIC(Rack_Murr_Node4_Instrum_TFF2.Node_Comm_Status) ,XIC(Rack_Murr_Node4_Instrum_TFF3.Node_Comm_Status) ,XIC(Rack_Murr_Node4_Instrum_TFF4.Node_Comm_Status) ,XIC(Rack_Murr_Node4_Instrum_TFF5.Node_Comm_Status) ]GSV(Module,RACK_MURR_NODE4_INSTRUM_TFF1,Mode,Rack_Murr_Node4_Instrum_TFF1.Inhibition)OR(Rack_Murr_Node4_Instrum_TFF1.Inhibition,4,Rack_Murr_Node4_Instrum_TFF1.Inhibition)SSV(Module,RACK_MURR_NODE4_INSTRUM_TFF1,Mode,Rack_Murr_Node4_Instrum_TFF1.Inhibition);
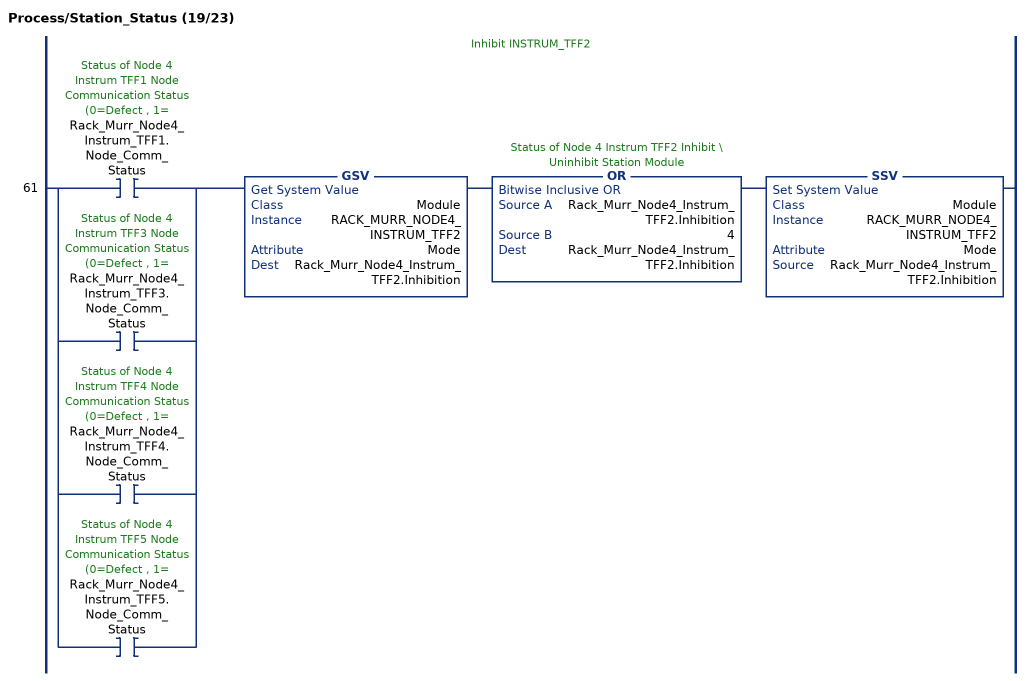
   // Inhibit INSTRUM_TFF2
   61: [XIC(Rack_Murr_Node4_Instrum_TFF1.Node_Comm_Status) ,XIC(Rack_Murr_Node4_Instrum_TFF3.Node_Comm_Status) ,XIC(Rack_Murr_Node4_Instrum_TFF4.Node_Comm_Status) ,XIC(Rack_Murr_Node4_Instrum_TFF5.Node_Comm_Status) ]GSV(Module,RACK_MURR_NODE4_INSTRUM_TFF2,Mode,Rack_Murr_Node4_Instrum_TFF2.Inhibition)OR(Rack_Murr_Node4_Instrum_TFF2.Inhibition,4,Rack_Murr_Node4_Instrum_TFF2.Inhibition)SSV(Module,RACK_MURR_NODE4_INSTRUM_TFF2,Mode,Rack_Murr_Node4_Instrum_TFF2.Inhibition);
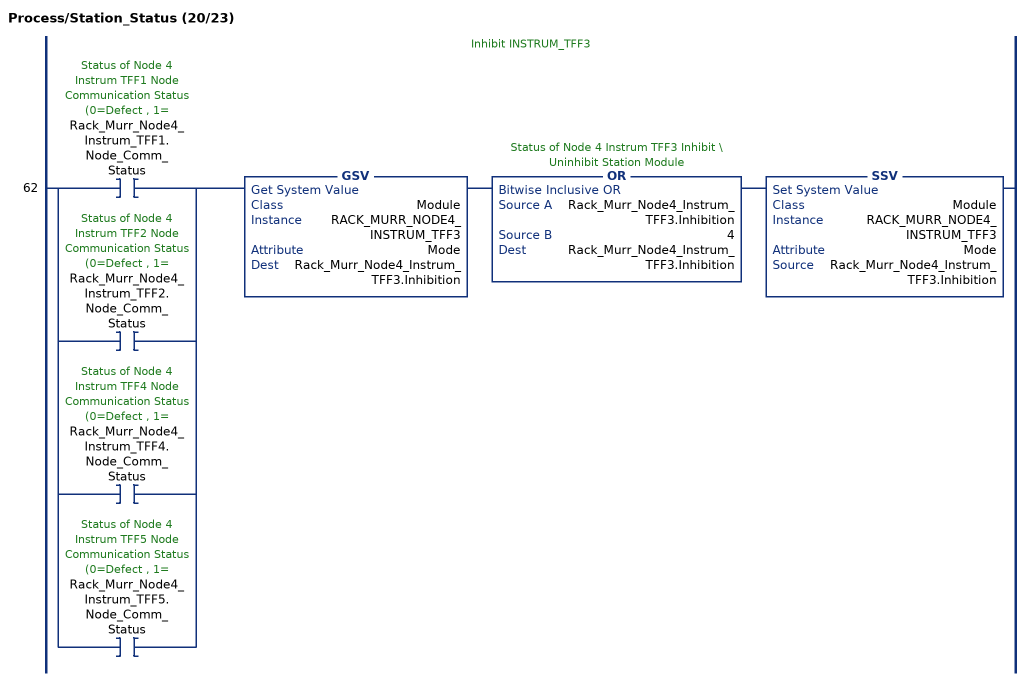
   // Inhibit INSTRUM_TFF3
   62: [XIC(Rack_Murr_Node4_Instrum_TFF1.Node_Comm_Status) ,XIC(Rack_Murr_Node4_Instrum_TFF2.Node_Comm_Status) ,XIC(Rack_Murr_Node4_Instrum_TFF4.Node_Comm_Status) ,XIC(Rack_Murr_Node4_Instrum_TFF5.Node_Comm_Status) ]GSV(Module,RACK_MURR_NODE4_INSTRUM_TFF3,Mode,Rack_Murr_Node4_Instrum_TFF3.Inhibition)OR(Rack_Murr_Node4_Instrum_TFF3.Inhibition,4,Rack_Murr_Node4_Instrum_TFF3.Inhibition)SSV(Module,RACK_MURR_NODE4_INSTRUM_TFF3,Mode,Rack_Murr_Node4_Instrum_TFF3.Inhibition);
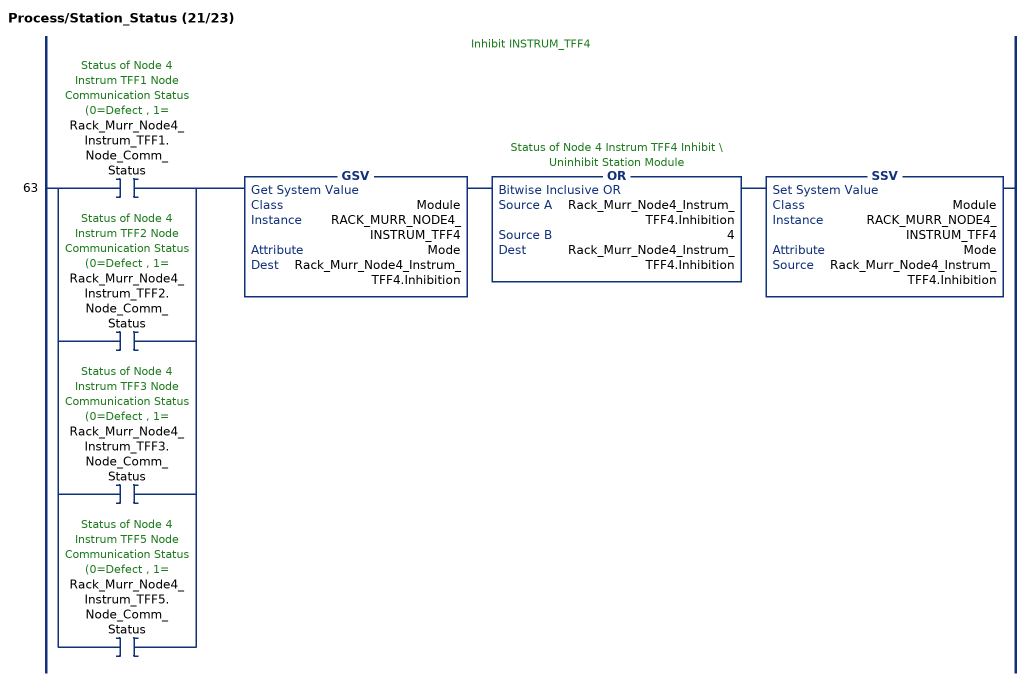
   // Inhibit INSTRUM_TFF4
   63: [XIC(Rack_Murr_Node4_Instrum_TFF1.Node_Comm_Status) ,XIC(Rack_Murr_Node4_Instrum_TFF2.Node_Comm_Status) ,XIC(Rack_Murr_Node4_Instrum_TFF3.Node_Comm_Status) ,XIC(Rack_Murr_Node4_Instrum_TFF5.Node_Comm_Status) ]GSV(Module,RACK_MURR_NODE4_INSTRUM_TFF4,Mode,Rack_Murr_Node4_Instrum_TFF4.Inhibition)OR(Rack_Murr_Node4_Instrum_TFF4.Inhibition,4,Rack_Murr_Node4_Instrum_TFF4.Inhibition)SSV(Module,RACK_MURR_NODE4_INSTRUM_TFF4,Mode,Rack_Murr_Node4_Instrum_TFF4.Inhibition);
